Fanuc KAREL source: KA00047.KL

PROGRAM KA00047
%NOLOCKGROUP
VAR
  SRC: STRING[80]
  DST: ARRAY[2] OF BYTE
BEGIN
  SRC = 'A'
  DST[1] = SRC
END KA00047
